(* IEC 61131-3 sources: plc_generation_empirical_study/datasets_50/tasks/C06_M02_bounded_up_down_counter, 2 files *)

(* ---- interface.st ---- *)
FUNCTION_BLOCK C06_M02_bounded_up_down_counter
VAR_INPUT
    AddItem : BOOL;
    RemoveItem : BOOL;
    Reset : BOOL;
    Capacity : INT;
END_VAR
VAR_OUTPUT
    Count : INT;
    Empty : BOOL;
    Full : BOOL;
    Conflict : BOOL;
END_VAR
END_FUNCTION_BLOCK

(* ---- reference.st ---- *)
FUNCTION_BLOCK C06_M02_bounded_up_down_counter
VAR_INPUT
    AddItem : BOOL;
    RemoveItem : BOOL;
    Reset : BOOL;
    Capacity : INT;
END_VAR
VAR_OUTPUT
    Count : INT;
    Empty : BOOL;
    Full : BOOL;
    Conflict : BOOL;
END_VAR
VAR
    PrevAdd : BOOL := FALSE;
    PrevRemove : BOOL := FALSE;
END_VAR

Conflict := FALSE;
IF Reset THEN
    Count := 0;
ELSIF AddItem AND (NOT PrevAdd) AND RemoveItem AND (NOT PrevRemove) THEN
    Conflict := TRUE;
ELSIF AddItem AND (NOT PrevAdd) AND (Count < Capacity) THEN
    Count := Count + 1;
ELSIF RemoveItem AND (NOT PrevRemove) AND (Count > 0) THEN
    Count := Count - 1;
END_IF;
Empty := Count = 0;
Full := Count >= Capacity;
PrevAdd := AddItem;
PrevRemove := RemoveItem;

END_FUNCTION_BLOCK
